(* IEC 61131-3 sources: plc-process-lib/src/POUs/Devices/FB_DigitalInput, 8 files *)

(* ---- FB_DigitalInput.decl.st ---- *)
// Назначение: дискретный вход: инверсия (НЗ-контакт), задержки включения и отключения (FB_Delay),
//             подмена значения с ограничением по времени, отказ канала со значением по eFailValue,
//             тревога по состоянию и тревога отказа канала. Режимы: Auto — измерение, Manual —
//             подмена, OutOfService; Local нет. Наследует FB_DeviceBase: тело — нормативный порядок
//             цикла.
// Автор:      kr0nsch
// Версия:     0.1.0
// Документ:   docs/fb/FB_DigitalInput.md
FUNCTION_BLOCK FB_DigitalInput EXTENDS FB_DeviceBase
VAR_INPUT
    xIn           : BOOL;            // сигнал канала
    xChannelFault : BOOL;            // диагностика обрыва/КЗ (NAMUR-датчики, модуль), ошибка обмена
END_VAR
VAR_IN_OUT
    stCmd : ST_DigitalInputCmd;      // команды HMI/SCADA (GVL_Hmi.st<TAG>Cmd)
END_VAR
VAR_IN_OUT CONSTANT
    stCfg : ST_DigitalInputCfg;      // параметры (GVL_Persist.st<TAG>Cfg), только чтение
END_VAR
VAR_OUTPUT
    xValue : BOOL;                   // значение для логики
    xValid : BOOL;                   // нет отказа канала (или подмена), Cfg была корректна, не OOS
    stSts  : ST_DigitalInputSts;     // состояние для HMI/SCADA
END_VAR
VAR
    stCfgLkg   : ST_DigitalInputCfg; // последняя корректная конфигурация (LKG)
    fbDebounce : FB_Delay;           // задержки включения и отключения
    fbSubst    : FB_Delay;           // длительность подмены (tSubstMax)
    xGood      : BOOL;               // значение после задержек; при отказе канала — значение отказа (DI-2)
    xDelayInit : BOOL := TRUE;       // задержки ещё не предустановлены (до первого вызова с корректной Cfg)
END_VAR
VAR_TEMP
    eRes      : E_CmdResult;         // результат ProcessMode
    xRaw      : BOOL;                // сигнал после инверсии, до задержек
    xFaultAct : BOOL;                // отказ канала учитывается (не OutOfService)
    xAlmCond  : BOOL;                // условие тревоги State
    rAlmValue : REAL;                // значение для событий тревог: 0.0 / 1.0
    wLowBits  : WORD;                // младший байт wStatus
    eDevSt    : E_Ne107Status;       // вклад логики устройства в NE 107
END_VAR

(* ---- CheckConfig.method.decl.st ---- *)
// Проверка конфигурации: биты wCfgErr дискретного входа (карта — docs/fb/FB_DigitalInput.md). Только
// считает, ничего не меняет
METHOD PROTECTED CheckConfig : WORD
VAR_IN_OUT CONSTANT
    stCfgIn : ST_DigitalInputCfg;   // проверяемая конфигурация
END_VAR
VAR
    wErr : WORD;                    // непройденные проверки
END_VAR

(* ---- CheckConfig.method.impl.st ---- *)
IF NOT (stCfgIn.eFailValue = E_DiFailValue.HoldLast OR stCfgIn.eFailValue = E_DiFailValue.ForceFalse
        OR stCfgIn.eFailValue = E_DiFailValue.ForceTrue)
THEN
    wErr := wErr OR GVL_Const.DI_CFG_FAIL_VALUE;
END_IF
IF NOT CheckAlarmCfg(astCfg := stCfgIn.astAlarm) THEN
    wErr := wErr OR GVL_Const.DI_CFG_ALARM;
END_IF
CheckConfig := wErr;

(* ---- FB_DigitalInput.impl.st ---- *)
// 0. Первый вызов (до ProcessMode): тип, число слотов тревог; режим «Измерение» в памяти режима,
//    подмена (Manual) даёт CheckFunction
IF xFirstCall THEN
    uiAlarmCount := GVL_Const.DI_ALARM_COUNT;
    eDevType := E_DeviceType.DigitalInput;
    xManualIsCheck := TRUE;
    stModeMem.eRemoteMode := E_DeviceMode.Auto;
END_IF

// 1. Время
BeginCycle();

// 2. Конфигурация (LKG): дальше логика читает только stCfgLkg
IF AcceptCfg(wErr := CheckConfig(stCfgIn := stCfg)) THEN
    stCfgLkg := stCfg;
END_IF

// 3. Reset: фиксируемых отказов нет (отказ канала снимается сам), результат команды — Accepted;
//    квитирование выполнит RunAlarms
IF xResetReq OR stCmd.stCommon.xReset THEN
    SetCmdResult(eResult := E_CmdResult.Accepted);
END_IF

// 4. Режим: Local нет, OutOfService разрешён всегда; память режима — stModeMem (A-06)
eRes := ProcessMode(xLocalSel := FALSE, xLocalSupported := FALSE, xOosAllowed := TRUE,
                    stCmd := stCmd.stCommon, stRetain := stModeMem);
IF eRes <> E_CmdResult.None THEN
    SetCmdResult(eResult := eRes);
END_IF

// 5. Подмена ограничена по времени: Manual длится tSubstMax — возврат в Auto (SubstExpired), как у AI.
//    Preset — чтобы новый запрос подмены в следующем вызове отсчитал tSubstMax заново
fbSubst(xIn := (eMode = E_DeviceMode.Manual) AND (stCfgLkg.tSubstMax > T#0S), tOnDelay := stCfgLkg.tSubstMax,
        itfTime := itfTimeAct);
IF fbSubst.xOut THEN
    SwitchRemoteMode(eNew := E_DeviceMode.Auto, stRetain := stModeMem);
    fbSubst.Preset(xValue := FALSE);
    SetCmdResult(eResult := E_CmdResult.SubstExpired);
END_IF

// 6. Сигнал: инверсия до задержек. При отказе канала сигнал не верен: задержки стоят на значении отказа
//    (HoldLast — значение до отказа, ForceFalse/ForceTrue — значение по eFailValue) и после возврата канала
//    отсчитываются от него заново: значение отказа снимается только через задержку, без провала защитного
//    сигнала (DI-2). В первом вызове с корректной Cfg значение берётся без задержки (DI-1): не в первом вызове
//    вообще — до корректной Cfg инверсия взята из умолчаний, и НЗ-контакт прошёл бы через задержку с неверной
//    полярностью
xRaw := xIn XOR stCfgLkg.xInvert;
IF xDelayInit AND xCfgEverOk THEN
    xGood := xRaw AND NOT xChannelFault;
    fbDebounce.Preset(xValue := xGood);
    xDelayInit := FALSE;
END_IF
IF xChannelFault THEN
    // значение отказа: HoldLast — прежнее, ForceTrue — TRUE, ForceFalse — FALSE (eFailValue проверен CheckConfig)
    xGood := (xGood AND stCfgLkg.eFailValue = E_DiFailValue.HoldLast) OR stCfgLkg.eFailValue = E_DiFailValue.ForceTrue;
    fbDebounce.Preset(xValue := xGood);
ELSE
    fbDebounce(xIn := xRaw, tOnDelay := stCfgLkg.tOnDelay, tOffDelay := stCfgLkg.tOffDelay, itfTime := itfTimeAct);
    xGood := fbDebounce.xOut;
END_IF

// Выбор значения по режиму и состоянию канала
xFaultAct := xChannelFault AND eMode <> E_DeviceMode.OutOfService;
SelectValue(xSubst := stCmd.xSubstValue);

// Слежение: пока значением управляет не оператор, ФБ пишет текущее значение в поле подмены —
// переход в подмену без рывка
IF eMode <> E_DeviceMode.Manual THEN
    stCmd.xSubstValue := xValue;
END_IF

// 7. Тревоги (слоты E_DiAlarm): State подавляется при отказе канала — отказ показывает слот Failure
//    (без дублирования по ISA-18.2). Значение события — xValue как 0.0 / 1.0
xAlmCond := xValue = stCfgLkg.xAlarmOnTrue;
rAlmValue := SEL(xValue, 0.0, 1.0);
axAlmCond[E_DiAlarm.State] := xAlmCond;
axAlmCond[E_DiAlarm.Failure] := xChannelFault;
axAlmSuppress[E_DiAlarm.State] := xChannelFault;
axAlmSuppress[E_DiAlarm.Failure] := FALSE;
arAlmValue[E_DiAlarm.State] := rAlmValue;
arAlmValue[E_DiAlarm.Failure] := rAlmValue;
RunAlarms(udiIdBase := stCfgLkg.udiAlarmIdBase, stCmd := stCmd.stCommon, astCfg := stCfgLkg.astAlarm);

// 8. Состояние; биты отсчёта задержек — пока канал исправен
wLowBits := SEL(xValue, 0, GVL_Const.DI_STS_VALUE) OR SEL(xRaw, 0, GVL_Const.DI_STS_RAW)
            OR SEL(fbDebounce.xTimingOn AND NOT xChannelFault, 0, GVL_Const.DI_STS_TIMING_ON)
            OR SEL(fbDebounce.xTimingOff AND NOT xChannelFault, 0, GVL_Const.DI_STS_TIMING_OFF)
            OR SEL(xChannelFault, 0, GVL_Const.DI_STS_CHANNEL_FAULT)
            OR SEL(xAlmCond, 0, GVL_Const.DI_STS_ALARM_COND);
IF xFaultAct THEN
    eDevSt := E_Ne107Status.Failure;
ELSE
    eDevSt := E_Ne107Status.Good;
END_IF
stSts.uiSubstRemain_s := SubstRemainSec();
FinishCycle(eDevStatus := eDevSt, xAvailableDev := xValid, wLow := wLowBits,
            wFaultBits := SEL(xFaultAct, 0, GVL_Const.DI_FLT_CHANNEL), wWarnBits := 0,
            stCommon := stSts.stCommon);

(* ---- SelectValue.method.decl.st ---- *)
// Шаг 6 цикла: значение для логики xValue и xValid (контракт 12.3, таблица 2.6). Нет корректной Cfg —
// FALSE; OutOfService — удержание; Manual — подмена без задержек; отказ канала — значение отказа xGood
// (тело выставляет его по eFailValue: HoldLast — значение до отказа), xValid = FALSE. Значение подмены
// приходит параметром: метод не читает VAR_IN_OUT (R2)
METHOD PROTECTED SelectValue
VAR_INPUT
    xSubst : BOOL;   // значение подмены stCmd.xSubstValue
END_VAR

(* ---- SelectValue.method.impl.st ---- *)
IF NOT xCfgEverOk THEN
    // безопасное значение: корректной Cfg ещё не было
    xValue := FALSE;
    xValid := FALSE;
ELSIF eMode = E_DeviceMode.OutOfService THEN
    // значение удерживается
    xValid := FALSE;
ELSIF eMode = E_DeviceMode.Manual THEN
    xValue := xSubst;
    xValid := TRUE;
ELSIF xChannelFault THEN
    // значение отказа: тело выставило xGood по eFailValue (HoldLast — значение до отказа)
    xValue := xGood;
    xValid := FALSE;
ELSE
    xValue := xGood;
    xValid := TRUE;
END_IF

(* ---- SubstRemainSec.method.decl.st ---- *)
// Остаток подмены для stSts.uiSubstRemain_s: целые секунды с округлением вверх (пока подмена идёт,
// остаток не 0), не больше UINT_MAX. 0 — подмены нет или её срок не ограничен (tSubstMax = T#0S)
METHOD PROTECTED SubstRemainSec : UINT
VAR
    lrRemain_s  : LREAL;   // до снятия подмены, с
    udiRemain_s : UDINT;   // то же, целых секунд
END_VAR

(* ---- SubstRemainSec.method.impl.st ---- *)
IF eMode = E_DeviceMode.Manual AND stCfgLkg.tSubstMax > T#0S THEN
    lrRemain_s := F_TimeToSec(tIn := fbSubst.tRemaining);
    udiRemain_s := LREAL_TO_UDINT(lrRemain_s);
    IF UDINT_TO_LREAL(udiRemain_s) < lrRemain_s THEN
        udiRemain_s := udiRemain_s + 1;
    END_IF
    SubstRemainSec := UDINT_TO_UINT(MIN(udiRemain_s, UINT_TO_UDINT(GVL_Const.UINT_MAX)));
ELSE
    SubstRemainSec := 0;
END_IF
